ABB RAPID module: TCP_Hfeli.mod

MODULE TCP_Hfeli
	! Points are read in order of declaration.
  ! Please do not change the order of points!

  LOCAL PERS robtarget pTCP_Point1:=[[577.3022,0.1874072,383.2325],[0.178669765591621,-0.00116579560562968,0.98390805721283,-0.000844044843688607],[0,-1,-1,0],[9E+09,9E+09,9E+09,9E+09,9E+09,9E+09]];
	LOCAL PERS robtarget pTCP_Point2:=[[521.1808,76.69171,369.1685],[0.158674284815788,-0.585275530815125,0.790488243103027,-0.0860425606369972],[0,-1,-1,0],[9E+09,9E+09,9E+09,9E+09,9E+09,9E+09]];
	LOCAL PERS robtarget pTCP_Point3:=[[490.0894,-95.00866,347.4818],[0.359917670488358,0.423246383666992,0.772478580474854,0.30756875872612],[-1,1,-1,0],[9E+09,9E+09,9E+09,9E+09,9E+09,9E+09]];
	LOCAL PERS robtarget pTCP_Point4:=[[470.696,5.853047,383.0463],[0.0190307293087244,-0.988126754760742,0.077323243021965,0.131394192576408],[0,0,-2,0],[9E+09,9E+09,9E+09,9E+09,9E+09,9E+09]];

ENDMODULE
